VISUALIZATION FP_Test  // 2x2
VAR_IN_OUT
	bTest : BOOL;
END_VAR
END_VISUALIZATION

(* stored: Version 1.1.0.1
   Visu FP_Test: Id {0daa2f4a-98c7-4ce0-873c-726b003f9f24} *)
